Fanuc KAREL source: kt00060.KL

-- PROVISIONAL review KL for V1013-1; original PC SHA256 39437fe439a9f84079a0223278fbdd85f92a6c79f29680a43f64fcd8c7b02308
-- Incomplete behavior may be omitted. Consult companion uncertainty JSON. Do not deploy.
PROGRAM KT00060
%NOLOCKGROUP
VAR
  R2 : REAL
  OUT : REAL
-- UNRESOLVED_DECL H1 type=002017
BEGIN
  -- UNRESOLVED_PC offsets 5-19; opcodes 2E,22,9D,33,B4
  -- UNRESOLVED_PC offsets 24-35; opcodes 2E,23
  -- UNRESOLVED_PC offsets 40-65; opcodes 22,9D,33,B3,21,29,64,29,6A,23
  -- UNRESOLVED_PC offsets 70-74; opcodes 7F
END KT00060
